(* IEC 61131-3 sources: PLC-Static-Analysis/modules/plc-rules/src/test/resources/PLCA-Q010, 2 files *)

(* ---- compliant.st ---- *)
FUNCTION F_Ok : INT
VAR_INPUT
    bMode : BOOL;
    n : INT;
END_VAR
VAR
    nPick : INT;
    nInit : INT := 5;
    nBoth : INT;
    nCase : INT;
    nRep : INT;
    nOut : INT;
    nAdr : INT;
    p : POINTER TO INT;
    stData : ST_Data;
END_VAR
IF bMode THEN
    nBoth := 1;
ELSE
    nBoth := 2;
END_IF
CASE n OF
    1: nCase := 1;
    ELSE nCase := 0;
END_CASE
REPEAT
    nRep := 1;
UNTIL TRUE
END_REPEAT
IF n < 0 THEN
    RETURN;
ELSE
    nPick := n;
END_IF
F_Out(n := n, nOut => nOut);
p := ADR(nAdr);
F_Ok := nPick + nInit + nBoth + nCase + nOut + nAdr + stData.a;
END_FUNCTION

FUNCTION F_Out : BOOL
VAR_INPUT
    n : INT;
END_VAR
VAR_OUTPUT
    nOut : INT;
END_VAR
nOut := n;
END_FUNCTION

TYPE ST_Data :
STRUCT
    a : INT;
END_STRUCT
END_TYPE

FUNCTION_BLOCK FB_Static
VAR
    nCount : INT;
END_VAR
nCount := nCount + 1;
END_FUNCTION_BLOCK

(* ---- noncompliant.st ---- *)
FUNCTION F_Sum : INT
VAR_INPUT
    a : ARRAY[0..3] OF INT;
    bMode : BOOL;
END_VAR
VAR
    i : INT;
    nSum : INT;
    nLast : INT;
    nPick : INT;
    nOnce : INT;
END_VAR
FOR i := 0 TO 3 DO
    nSum := nSum + a[i]; // accumulator on the zero default: not reported
END_FOR
IF bMode THEN
    nPick := 1;
END_IF
F_Sum := nPick; // PLCA-Q010
F_Sum := F_Sum + nLast; // PLCA-Q010
WHILE i > 0 DO
    nOnce := 1;
    i := i - 1;
END_WHILE
F_Sum := F_Sum + nOnce; // PLCA-Q010
END_FUNCTION

FUNCTION_BLOCK FB_Temp
VAR_TEMP
    nTmp : INT;
END_VAR
VAR
    nStatic : INT;
END_VAR
nStatic := nStatic + nTmp; // PLCA-Q010
END_FUNCTION_BLOCK

FUNCTION F_Result : INT
F_Result := F_Result + 1; // self-update: not reported
END_FUNCTION
